FUNCTION F_TxtBatCmd : WSTRING(31)
VAR_INPUT
	i_e		: E_BatCmd;
END_VAR

CASE i_e OF
	E_BatCmd.None:		F_TxtBatCmd := "없음";
	E_BatCmd.Close:		F_TxtBatCmd := "배터리 투입";
	E_BatCmd.Open:		F_TxtBatCmd := "배터리 개방";
	E_BatCmd.EStop:		F_TxtBatCmd := "배터리 비상정지";
	E_BatCmd.Reset:		F_TxtBatCmd := "배터리 Reset";
ELSE
	F_TxtBatCmd := "?";
END_CASE

END_FUNCTION

(* stored: Version 1.1.0.1, ProductVersion 3.1.4024.15
   POU F_TxtBatCmd: Id {c64104e3-b7a8-4e0e-8a3e-bfb1549ef29d}, SpecialFunc None *)
